(* IEC 61131-3 sources: AyCD/codesys/src/GVLs, 3 files *)

(* ---- GVL_COMMS.st ---- *)
(*
 * GVL_COMMS - Buffers UDP y estructuras de comunicación.
 * Las estructuras son escritas/leídas por COM_UDP_RX y COM_UDP_TX.
 *)
VAR_GLOBAL
    // Estructura recibida de Simulink (lo que el PLC lee)
    udp_from_sim       : T_UDP_TX_FROM_SIM;

    // Estructura enviada a Simulink (lo que el PLC escribe)
    udp_to_sim         : T_UDP_RX_TO_SIM;

    // Estado conexión
    udp_rx_socket      : DINT := -1;
    udp_tx_socket      : DINT := -1;
    udp_rx_ok          : BOOL := FALSE;
    udp_tx_ok          : BOOL := FALSE;
    udp_rx_count       : UDINT := 0;        // contador paquetes recibidos
    udp_tx_count       : UDINT := 0;        // contador paquetes enviados
    udp_rx_err         : DINT := 0;
    udp_tx_err         : DINT := 0;
END_VAR

(* ---- GVL_PARAMS.st ---- *)
(*
 * GVL_PARAMS - Constantes físicas y de configuración
 * Espejo de simulink/init_plant_parameters.m
 *)
VAR_GLOBAL CONSTANT
    // === Tiempos de muestreo ===
    Ts0                : LREAL := 0.02;          // [s] Nivel 0 (seguridad)
    Ts1                : LREAL := 0.02;          // [s] Nivel 1 (supervisor)
    Ts2                : LREAL := 0.001;         // [s] Nivel 2 (torque)

    // === Constantes universales ===
    g                  : LREAL := 9.80665;       // [m/s^2] gravedad
    Yt0                : LREAL := 45.0;          // [m] altura poleas
    Ysb                : LREAL := 5.0;           // [m] despeje sobre testera

    // === Masas y containers ===
    Ms                 : LREAL := 15000.0;       // [kg] spreader + headblock
    Mc_max             : LREAL := 50000.0;       // [kg] container máximo
    Mc_min             : LREAL := 2000.0;        // [kg] container vacío
    Hc                 : LREAL := 2.59;          // [m] altura container ISO
    Wc                 : LREAL := 2.44;          // [m] ancho container ISO

    // === Izaje (hoist) ===
    rhd                : LREAL := 0.75;          // [m] radio tambor izaje
    ih                 : LREAL := 22.0;          // relación transmisión izaje
    yh_min             : LREAL := -20.0;         // [m] límite inferior
    yh_max             : LREAL := 40.0;          // [m] límite superior
    vh_max             : LREAL := 3.0;           // [m/s] vel max sin carga
    vh_nom             : LREAL := 1.5;           // [m/s] vel nominal
    ah_max             : LREAL := 0.75;          // [m/s^2] aceleración max
    P_nom              : LREAL := 956150.0;      // [W] potencia nominal

    // === Carro (trolley) ===
    Mt                 : LREAL := 30000.0;       // [kg] masa carro
    rtd                : LREAL := 0.50;          // [m] radio tambor carro
    it                 : LREAL := 30.0;          // relación transmisión carro
    xt_min             : LREAL := -30.0;         // [m] límite mínimo
    xt_max             : LREAL := 50.0;          // [m] límite máximo
    vt_max             : LREAL := 4.0;           // [m/s] vel max
    at_max             : LREAL := 0.80;          // [m/s^2] acel max

    // === Watchdog y comunicación ===
    periodo_pulsos     : LREAL := 0.1;           // [s] pulso heartbeat cada 100 ms
    timeout_wd         : LREAL := 0.3;           // [s] timeout watchdog
    counter_limit      : DINT  := 15;            // ciclos (= timeout/Ts0)

    // === Modo manual ===
    dead_zone          : LREAL := 0.1;           // zona muerta joystick

    // === Perfil ===
    N_xt               : INT   := 33;            // cantidad de columnas perfil
    alt_borde          : LREAL := 2.8;           // [m] altura borde muelle

    // === UDP ===
    UDP_PORT_RX        : UINT  := 25000;         // PLC escucha (Sim TX)
    UDP_PORT_TX        : UINT  := 25001;         // PLC envía (Sim RX)
    UDP_REMOTE_IP      : STRING := '127.0.0.1';

    // === Tamaños paquetes ===
    UDP_RX_SIZE        : UDINT := 248;           // bytes paquete TX_FROM_SIM
    UDP_TX_SIZE        : UDINT := 424;           // bytes paquete RX_TO_SIM
END_VAR

(* ---- GVL_PROCESS.st ---- *)
(*
 * GVL_PROCESS - Señales compartidas entre L0 (CONTROL_SEGURIDAD)
 * y L1 (CONTROL_SUPERVISOR). Solo un POU escribe cada variable.
 *)
VAR_GLOBAL
    // === Escrito por L1, leído por L0 ===
    heartbeat_L1       : INT  := 0;          // pulso watchdog (toggle por ciclo L1)
    m_container_L1     : LREAL := 0.0;       // masa container estimada [kg]
    modo_muerto_L1     : BOOL := FALSE;      // flag modo muerto desde supervisor

    // === Escrito por L0, leído por L1 ===
    FALLA_GLOBAL       : BOOL := FALSE;      // cualquier falla activa
    FALLA_MAN_L0       : BOOL := FALSE;      // emergencia manual
    FALLA_WD_L0        : BOOL := FALSE;      // timeout watchdog
    FALLA_SV_L0        : BOOL := FALSE;      // sobrevelocidad
    FALLA_CARRO_DER_L0 : BOOL := FALSE;
    FALLA_CARRO_IZQ_L0 : BOOL := FALSE;
    FALLA_CARRO_SV_L0  : BOOL := FALSE;
    FALLA_IZAJE_INF_L0 : BOOL := FALSE;
    FALLA_IZAJE_SUP_L0 : BOOL := FALSE;
    FALLA_IZAJE_SV_L0  : BOOL := FALSE;
    RECUPERAR_L0       : BOOL := FALSE;      // pedido de recuperación a L1
    vh_lim_L0          : LREAL := 3.0;       // velocidad izaje límite dinámica

    // === Salidas de frenos (ambos niveles) ===
    BRK_h_N0           : INT  := 0;          // 0 = liberado, 1 = frenado
    BRK_t_N0           : INT  := 0;
    BRK_h_N1           : INT  := 0;
    BRK_t_N1           : INT  := 0;

    // === Salidas supervisor ===
    TLK_OUT            : INT  := 0;
    vx_suave           : LREAL := 0.0;
    vy_suave           : LREAL := 0.0;
    i_sel_OUT          : INT  := 0;
    recuperacion_OUT   : BOOL := FALSE;
    yc0_vec_OUT        : ARRAY[1..33] OF LREAL;
END_VAR
